(*
| This function block is based on a _`statemachine` concept which is described in the following.
| The statemachine is based on several states.
| The proceeding always begins in the first state.
| If the last state is left, the execution restarts in the first state.
| There are so many more information necessary to describe the statemachine concept in detail.
| But as this is just a sample text to show the inline hyperlinks, we want to leave out the details.
| A rough description should be enough for the sample demonstration.
| 
| Some sample text to get some text in between.
| Some sample text to get some text in between.
| Some sample text to get some text in between.
| Some sample text to get some text in between.
| Some sample text to get some text in between.
| Some sample text to get some text in between.
| 
| Furthermore, the function block is based on another concept. This is called XY.
| It is always necessary to respect the demands of this concept.
| Especially, as it is deeply interwoven with the statemachine concept.
| Therefore, you definitely need to understand the statemachine concept first.
| Afterwards, you might understand the XY concept.
| For more information about this, see the description of the `statemachine`_.
| By clicking on this link, the Library Manager will jump to the beginning of the first paragraph where the statemachine concept is described.. 

*)

FUNCTION_BLOCK FB_Libdoc_InlineHyperlinks
VAR_INPUT
    nVarA : INT;
    nVarB : INT;
END_VAR
VAR_OUTPUT
    nSum : INT;
END_VAR
VAR
END_VAR

END_FUNCTION_BLOCK

(* stored: Version 1.1.0.1, ProductVersion 3.1.4024.0
   POU FB_Libdoc_InlineHyperlinks: Id {601f44cb-a066-41cb-8892-2ccc238675fc}, SpecialFunc None *)
